(* IEC 61131-3 sources: STAR-PLC-Agent/results/raw/codex_matrix_resume_20261114/codex_terra/SELF003/formal/attempt_0001, 1 file *)

(* ---- candidate.st ---- *)
FUNCTION_BLOCK FB_Task
VAR_INPUT
    Start : BOOL;
    Stop : BOOL;
    EStopNC : BOOL;
    Reset : BOOL;
END_VAR
VAR_OUTPUT
    Run : BOOL := FALSE;
    ResetRequired : BOOL := TRUE;
END_VAR

IF NOT EStopNC THEN
    ResetRequired := TRUE;
    Run := FALSE;
ELSIF ResetRequired THEN
    Run := FALSE;
    IF Reset AND NOT Start AND NOT Stop THEN
        ResetRequired := FALSE;
    END_IF;
ELSIF Stop THEN
    Run := FALSE;
ELSIF Start THEN
    Run := TRUE;
END_IF;
END_FUNCTION_BLOCK
